(* IEC 61131-3 sources: Simulierte-Foerderanlagensteuerung/plc/simulation, 3 files *)

(* ---- GVL_Simulation.st ---- *)
(* ============================================================================
   GVL_Simulation.st
   Globale Variablen der Anlagensimulation (elektrisches/mechanisches Modell).

   ACHTUNG: Diese Variablen existieren NUR in der Simulation. Sie bilden das
   Verhalten von Schuetz, Motor, Motorschutz und Foerderband nach und erlauben
   eine gezielte Fehlerinjektion fuer Tests und Diagnose.
   ============================================================================ *)

VAR_GLOBAL
    (* --- Fehlerinjektion (nur Simulation) --- *)
    xSimInjectOverload            : BOOL;  (* Motorschutz nach T_OVERLOAD_TRIP ausloesen *)
    xSimInjectFeedbackOpen        : BOOL;  (* Rueckmeldung faellt aus (laeuft nicht an) *)
    xSimInjectFeedbackStuck       : BOOL;  (* Rueckmeldung haengt (stoppt nicht) *)
    xSimInjectJam                 : BOOL;  (* Band blockiert (Stau) *)
    xSimInjectSensorInconsistency : BOOL;  (* Auslaufsensor liefert Dauersignal *)
    xSimGenerateWorkpieces        : BOOL;  (* Werkstuecke automatisch erzeugen *)
    xSimResetCount                : BOOL;  (* Werkstueckzaehler ruecksetzen *)

    (* --- Simulations-Anzeigewerte --- *)
    xSimOverloadTrip  : BOOL;  (* Motorschutz F2 ausgeloest *)
    xSimContactor     : BOOL;  (* Schuetz K1 angezogen *)
    xSimMotorRunning  : BOOL;  (* Motor laeuft (mechanisch) *)
END_VAR

(* ---- FB_BeltSimulation.st ---- *)
(* ============================================================================
   FB_BeltSimulation.st
   Mechanisches Modell des Foerderbands.

   - Das Band hat eine normierte Laenge von 0..100 %.
   - Werkstuecke werden in 5 Plaetzen gefuehrt (aPos; -1 = frei).
   - Bei laufendem Motor bewegen sich die Werkstuecke mit BELT_SPEED_PER_S.
   - Beim Durchlaufen der Zonen werden die Sensoren B1 (Einlauf) und B2 (Auslauf)
     gesetzt.
   - xInjectJam blockiert den Transport (Stau).
   - xInjectSensorInconsistency erzwingt ein dauerhaftes Auslaufsignal.
   ============================================================================ *)

FUNCTION_BLOCK FB_BeltSimulation
VAR_INPUT
    xMotorRunning              : BOOL;
    xGenerate                  : BOOL;   (* Werkstuecke automatisch erzeugen *)
    xInjectJam                 : BOOL;
    xInjectSensorInconsistency : BOOL;
END_VAR
VAR_OUTPUT
    xEntrySensor : BOOL;                 (* B1 *)
    xExitSensor  : BOOL;                 (* B2 *)
    aPos         : ARRAY[0..4] OF REAL;  (* Werkstueckpositionen in % *)
END_VAR
VAR
    i          : INT;
    xInitDone  : BOOL;
    xPlaced    : BOOL;
    rStep      : REAL;
    tonGen     : TON;
END_VAR

    (* --- Einmalige Initialisierung --- *)
    IF NOT xInitDone THEN
        FOR i := 0 TO 4 DO
            aPos[i] := -1.0;
        END_FOR;
        xInitDone := TRUE;
    END_IF;

    (* --- Werkstuecke periodisch erzeugen (nur wenn gewuenscht) --- *)
    tonGen(IN := NOT tonGen.Q, PT := WORKPIECE_INTERVAL);
    IF xGenerate AND tonGen.Q THEN
        xPlaced := FALSE;
        FOR i := 0 TO 4 DO
            IF (NOT xPlaced) AND (aPos[i] < 0.0) THEN
                aPos[i] := 0.0;
                xPlaced := TRUE;
            END_IF;
        END_FOR;
    END_IF;

    (* --- Transport --- *)
    rStep := BELT_SPEED_PER_S * CYCLE_TIME_S;
    FOR i := 0 TO 4 DO
        IF aPos[i] >= 0.0 THEN
            IF xMotorRunning THEN
                IF NOT xInjectJam THEN
                    aPos[i] := aPos[i] + rStep;
                ELSE
                    (* Blockade in Bandmitte: Werkstueck laeuft bis 50 % und bleibt stehen *)
                    IF aPos[i] < 50.0 THEN
                        aPos[i] := aPos[i] + rStep;
                        IF aPos[i] > 50.0 THEN
                            aPos[i] := 50.0;
                        END_IF;
                    END_IF;
                END_IF;
            END_IF;
            IF aPos[i] > 100.0 THEN
                aPos[i] := -1.0;   (* Werkstueck hat das Band verlassen *)
            END_IF;
        END_IF;
    END_FOR;

    (* --- Sensorauswertung (Zonen) ---------------------------------------
       Einlaufzone 0..6 %: ein von der Zufuehrung aufgesetztes Werkstueck
       loest B1 unmittelbar aus.
       Auslaufzone 94..100 %: B2 wird bis zum Bandende gehalten.        *)
    xEntrySensor := FALSE;
    xExitSensor := FALSE;
    FOR i := 0 TO 4 DO
        IF (aPos[i] >= 0.0) AND (aPos[i] <= 6.0) THEN
            xEntrySensor := TRUE;
        END_IF;
        IF (aPos[i] >= 94.0) AND (aPos[i] <= 100.0) THEN
            xExitSensor := TRUE;
        END_IF;
    END_FOR;

    (* --- Fehlerinjektion: dauerhaftes Auslaufsignal --- *)
    IF xInjectSensorInconsistency THEN
        xExitSensor := TRUE;
    END_IF;
END_FUNCTION_BLOCK

(* ---- FB_ContactorMotor.st ---- *)
(* ============================================================================
   FB_ContactorMotor.st
   Simulationsmodell des elektrischen Leistungsteils:

       Schütz K1  ->  Drehstrommotor M1
       Motorschutzrelais F2 (Überlast)
       Rückmeldung (Hilfskontakt)

   WICHTIG (Konzept Leistungskreis vs. Steuerkreis):
   Das Schütz zieht nur an, wenn die SPS-Ansteuerung EIN ist UND keine harte
   Schutzbedingung (Überlast, Not-Halt) ansteht. Damit wirkt der Schutz
   unabhängig von der Software - genau wie in einer realen Schützung.
   ============================================================================ *)

FUNCTION_BLOCK FB_ContactorMotor
VAR_INPUT
    xCoilCmd             : BOOL;   (* Ansteuerung von der SPS (K1-Spule) *)
    xEmergencyActive     : BOOL;   (* Not-Halt-Kette offen -> harte Abschaltung *)
    xInjectOverload      : BOOL;   (* Fehlerinjektion Überlast *)
    xInjectFeedbackOpen  : BOOL;   (* Fehlerinjektion: Rückmeldung faellt aus *)
    xInjectFeedbackStuck : BOOL;   (* Fehlerinjektion: Rückmeldung haengt *)
END_VAR
VAR_OUTPUT
    xContactorClosed : BOOL;   (* Schütz angezogen (Hauptkontakt) *)
    xMotorRunning    : BOOL;   (* Motor laeuft (mechanisch) *)
    xMotorFeedback   : BOOL;   (* Rueckmeldung an die SPS *)
    xOverloadTrip    : BOOL;   (* Motorschutz F2 ausgeloest *)
END_VAR
VAR
    tonPull     : TON;
    tonOverload : TON;
    xEnergize   : BOOL;
END_VAR

    (* --- Motorschutzrelais F2: Auslösung bei anhaltender Überlast --- *)
    tonOverload(IN := xInjectOverload AND xMotorRunning, PT := T_OVERLOAD_TRIP);
    IF tonOverload.Q THEN
        xOverloadTrip := TRUE;
    END_IF;
    (* Manuelle Rückstellung des Schutzrelais (Injektion entfernt) *)
    IF NOT xInjectOverload THEN
        xOverloadTrip := FALSE;
        tonOverload(IN := FALSE, PT := T_OVERLOAD_TRIP);
    END_IF;

    (* --- Schützspule: harte Verriegelung durch Motorschutz und Not-Halt --- *)
    xEnergize := xCoilCmd AND NOT xOverloadTrip AND NOT xEmergencyActive;
    tonPull(IN := xEnergize, PT := T_CONTACTOR_PULL);
    xContactorClosed := tonPull.Q;

    (* --- Motor und Rückmeldung --- *)
    xMotorRunning := xContactorClosed;
    xMotorFeedback := xContactorClosed;

    (* --- Fehlerinjektion Rückmeldung --- *)
    IF xInjectFeedbackOpen THEN
        xMotorFeedback := FALSE;
    END_IF;
    IF xInjectFeedbackStuck THEN
        xMotorFeedback := TRUE;
    END_IF;
END_FUNCTION_BLOCK
